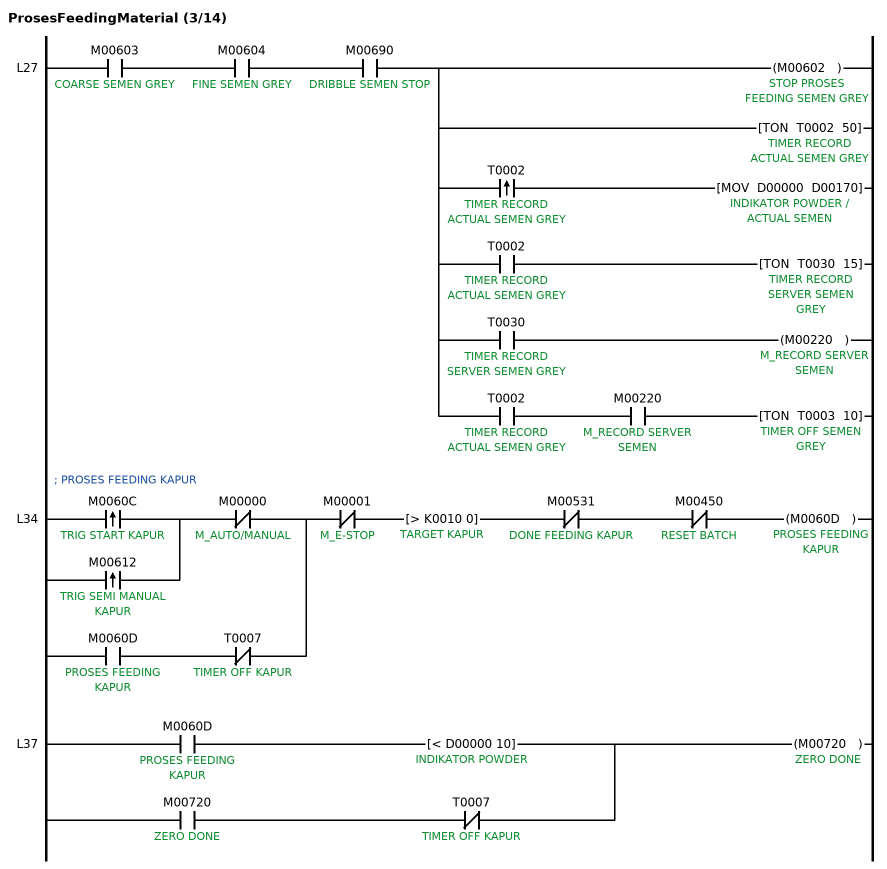
[picture p24: ProsesFeedingMaterial rungs L27-L37]
; L27
LOAD      M00603	// COARSE SEMEN GREY
AND       M00604	// FINE SEMEN GREY
AND       M00690	// DRIBBLE SEMEN STOP
OUT       M00602	// STOP PROSES FEEDING SEMEN GREY 
TON       T0002 50	// TIMER RECORD ACTUAL SEMEN GREY 
MPUSH
ANDP      T0002	// TIMER RECORD ACTUAL SEMEN GREY 
MOV       D00000 D00170	// INDIKATOR POWDER / ACTUAL SEMEN
MLOAD
AND       T0002	// TIMER RECORD ACTUAL SEMEN GREY 
TON       T0030 15	// TIMER RECORD SERVER SEMEN GREY
MLOAD
AND       T0030	// TIMER RECORD SERVER SEMEN GREY
OUT       M00220	// M_RECORD SERVER SEMEN
MPOP
AND       T0002	// TIMER RECORD ACTUAL SEMEN GREY 
AND       M00220	// M_RECORD SERVER SEMEN
TON       T0003 10	// TIMER OFF SEMEN GREY 
// PROSES FEEDING KAPUR
; L34
LOADP     M0060C	// TRIG START KAPUR
ORP       M00612	// TRIG SEMI MANUAL KAPUR 
AND NOT   M00000	// M_AUTO/MANUAL
LOAD      M0060D	// PROSES FEEDING KAPUR 
AND NOT   T0007	// TIMER OFF KAPUR
OR LOAD
AND NOT   M00001	// M_E-STOP
AND>      K0010 0	// TARGET KAPUR 
AND NOT   M00531	// DONE FEEDING KAPUR
AND NOT   M00450	// RESET BATCH
OUT       M0060D	// PROSES FEEDING KAPUR 
; L37
LOAD      M0060D	// PROSES FEEDING KAPUR 
AND<      D00000 10	// INDIKATOR POWDER
LOAD      M00720	// ZERO DONE
AND NOT   T0007	// TIMER OFF KAPUR
OR LOAD
OUT       M00720	// ZERO DONE

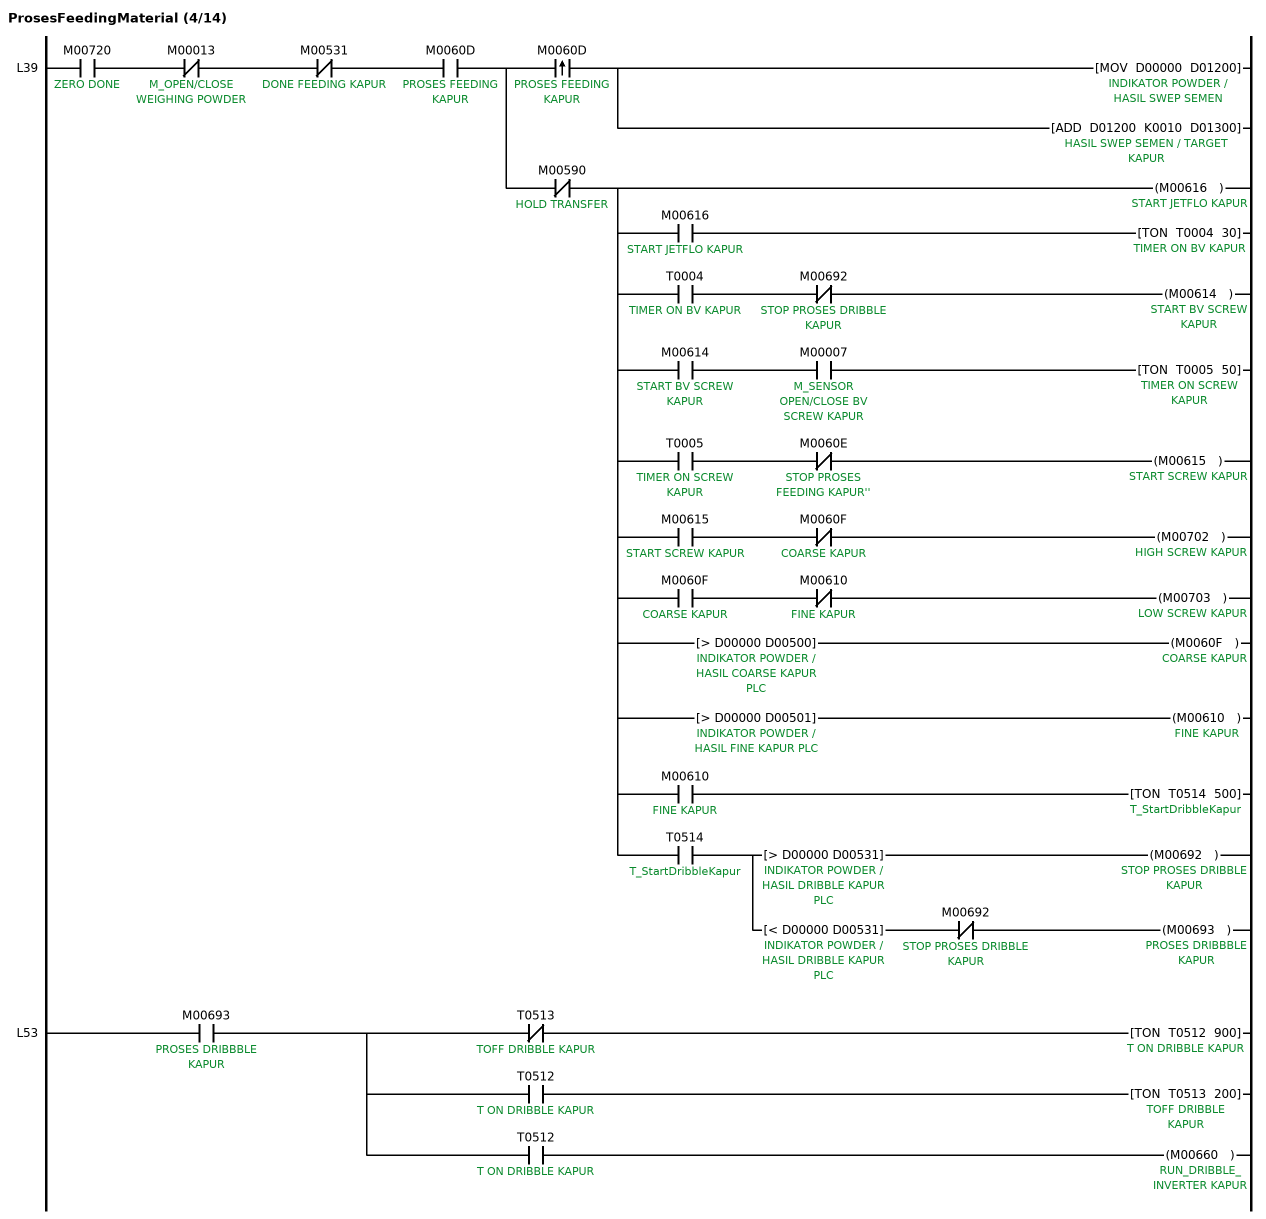
; L39
LOAD      M00720	// ZERO DONE
AND NOT   M00013	// M_OPEN/CLOSE WEIGHING POWDER
AND NOT   M00531	// DONE FEEDING KAPUR
AND       M0060D	// PROSES FEEDING KAPUR 
MPUSH
ANDP      M0060D	// PROSES FEEDING KAPUR 
MOV       D00000 D01200	// INDIKATOR POWDER / HASIL SWEP SEMEN
ADD       D01200 K0010 D01300	// HASIL SWEP SEMEN / TARGET KAPUR 
MPOP
AND NOT   M00590	// HOLD TRANSFER
OUT       M00616	// START JETFLO KAPUR
MPUSH
AND       M00616	// START JETFLO KAPUR
TON       T0004 30	// TIMER ON BV KAPUR
MLOAD
AND       T0004	// TIMER ON BV KAPUR
AND NOT   M00692	// STOP PROSES DRIBBLE KAPUR
OUT       M00614	// START BV SCREW KAPUR
MLOAD
AND       M00614	// START BV SCREW KAPUR
AND       M00007	// M_SENSOR OPEN/CLOSE BV SCREW KAPUR
TON       T0005 50	// TIMER ON SCREW KAPUR
MLOAD
AND       T0005	// TIMER ON SCREW KAPUR
AND NOT   M0060E	// STOP PROSES FEEDING KAPUR''
OUT       M00615	// START SCREW KAPUR
MLOAD
AND       M00615	// START SCREW KAPUR
AND NOT   M0060F	// COARSE KAPUR
OUT       M00702	// HIGH SCREW KAPUR
MLOAD
AND       M0060F	// COARSE KAPUR
AND NOT   M00610	// FINE KAPUR
OUT       M00703	// LOW SCREW KAPUR
MLOAD
AND>      D00000 D00500	// INDIKATOR POWDER / HASIL COARSE KAPUR PLC
OUT       M0060F	// COARSE KAPUR
MLOAD
AND>      D00000 D00501	// INDIKATOR POWDER / HASIL FINE KAPUR PLC 
OUT       M00610	// FINE KAPUR
MLOAD
AND       M00610	// FINE KAPUR
TON       T0514 500	// T_StartDribbleKapur
MPOP
AND       T0514	// T_StartDribbleKapur
MPUSH
AND>      D00000 D00531	// INDIKATOR POWDER / HASIL DRIBBLE KAPUR PLC 
OUT       M00692	// STOP PROSES DRIBBLE KAPUR
MPOP
AND<      D00000 D00531	// INDIKATOR POWDER / HASIL DRIBBLE KAPUR PLC 
AND NOT   M00692	// STOP PROSES DRIBBLE KAPUR
OUT       M00693	// PROSES DRIBBBLE KAPUR
; L53
LOAD      M00693	// PROSES DRIBBBLE KAPUR
MPUSH
AND NOT   T0513	// TOFF DRIBBLE KAPUR
TON       T0512 900	// T ON DRIBBLE KAPUR
MLOAD
AND       T0512	// T ON DRIBBLE KAPUR
TON       T0513 200	// TOFF DRIBBLE KAPUR
MPOP
AND       T0512	// T ON DRIBBLE KAPUR
OUT       M00660	// RUN_DRIBBLE_INVERTER KAPUR

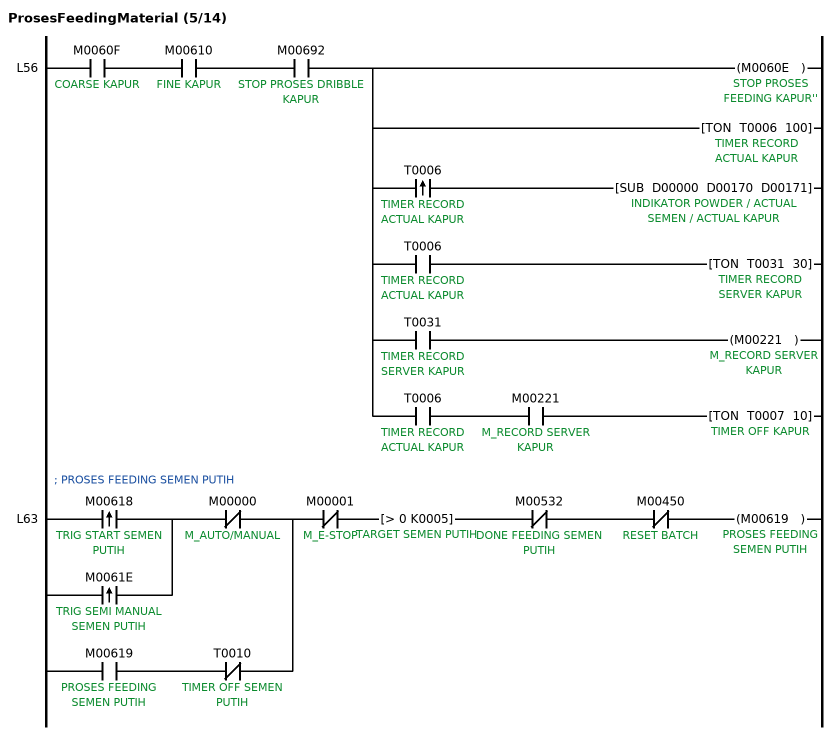
; L56
LOAD      M0060F	// COARSE KAPUR
AND       M00610	// FINE KAPUR
AND       M00692	// STOP PROSES DRIBBLE KAPUR
OUT       M0060E	// STOP PROSES FEEDING KAPUR''
TON       T0006 100	// TIMER RECORD ACTUAL KAPUR
MPUSH
ANDP      T0006	// TIMER RECORD ACTUAL KAPUR
SUB       D00000 D00170 D00171	// INDIKATOR POWDER / ACTUAL SEMEN / ACTUAL KAPUR
MLOAD
AND       T0006	// TIMER RECORD ACTUAL KAPUR
TON       T0031 30	// TIMER RECORD SERVER KAPUR
MLOAD
AND       T0031	// TIMER RECORD SERVER KAPUR
OUT       M00221	// M_RECORD SERVER KAPUR
MPOP
AND       T0006	// TIMER RECORD ACTUAL KAPUR
AND       M00221	// M_RECORD SERVER KAPUR
TON       T0007 10	// TIMER OFF KAPUR
// PROSES FEEDING SEMEN PUTIH
; L63
LOADP     M00618	// TRIG START SEMEN PUTIH
ORP       M0061E	// TRIG SEMI MANUAL SEMEN PUTIH
AND NOT   M00000	// M_AUTO/MANUAL
LOAD      M00619	// PROSES FEEDING SEMEN PUTIH 
AND NOT   T0010	// TIMER OFF SEMEN PUTIH
OR LOAD
AND NOT   M00001	// M_E-STOP
AND>      0 K0005	// TARGET SEMEN PUTIH
AND NOT   M00532	// DONE FEEDING SEMEN PUTIH 
AND NOT   M00450	// RESET BATCH
OUT       M00619	// PROSES FEEDING SEMEN PUTIH 

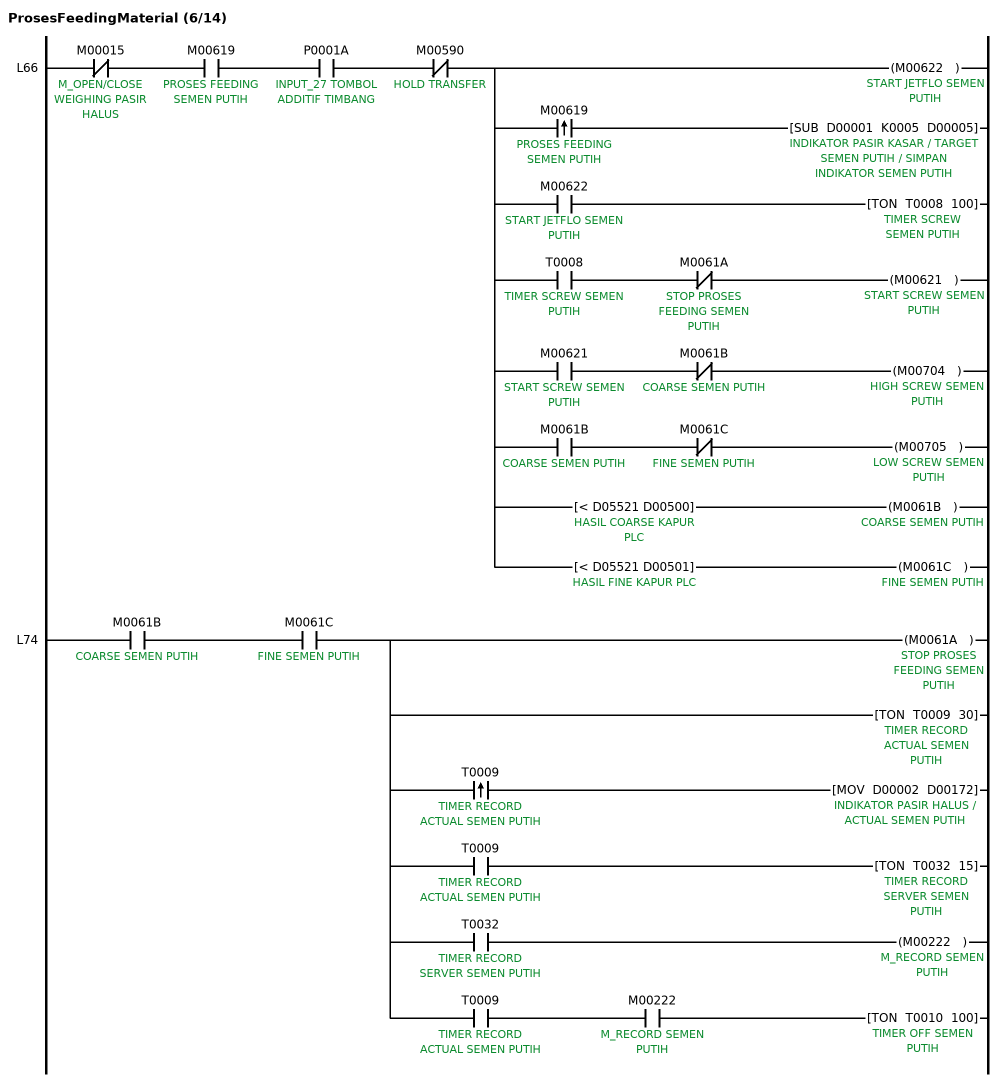
; L66
LOAD NOT  M00015	// M_OPEN/CLOSE WEIGHING PASIR HALUS 
AND       M00619	// PROSES FEEDING SEMEN PUTIH 
AND       P0001A	// INPUT_27 TOMBOL ADDITIF TIMBANG 
AND NOT   M00590	// HOLD TRANSFER
OUT       M00622	// START JETFLO SEMEN PUTIH
MPUSH
ANDP      M00619	// PROSES FEEDING SEMEN PUTIH 
SUB       D00001 K0005 D00005	// INDIKATOR PASIR KASAR / TARGET SEMEN PUTIH / SIMPAN INDIKATOR SEMEN PUTIH 
MLOAD
AND       M00622	// START JETFLO SEMEN PUTIH
TON       T0008 100	// TIMER SCREW SEMEN PUTIH
MLOAD
AND       T0008	// TIMER SCREW SEMEN PUTIH
AND NOT   M0061A	// STOP PROSES FEEDING SEMEN PUTIH
OUT       M00621	// START SCREW SEMEN PUTIH
MLOAD
AND       M00621	// START SCREW SEMEN PUTIH
AND NOT   M0061B	// COARSE SEMEN PUTIH
OUT       M00704	// HIGH SCREW SEMEN PUTIH 
MLOAD
AND       M0061B	// COARSE SEMEN PUTIH
AND NOT   M0061C	// FINE SEMEN PUTIH
OUT       M00705	// LOW SCREW SEMEN PUTIH 
MLOAD
AND<      D05521 D00500	// HASIL COARSE KAPUR PLC
OUT       M0061B	// COARSE SEMEN PUTIH
MPOP
AND<      D05521 D00501	// HASIL FINE KAPUR PLC 
OUT       M0061C	// FINE SEMEN PUTIH
; L74
LOAD      M0061B	// COARSE SEMEN PUTIH
AND       M0061C	// FINE SEMEN PUTIH
OUT       M0061A	// STOP PROSES FEEDING SEMEN PUTIH
TON       T0009 30	// TIMER RECORD ACTUAL SEMEN PUTIH
MPUSH
ANDP      T0009	// TIMER RECORD ACTUAL SEMEN PUTIH
MOV       D00002 D00172	// INDIKATOR PASIR HALUS / ACTUAL SEMEN PUTIH
MLOAD
AND       T0009	// TIMER RECORD ACTUAL SEMEN PUTIH
TON       T0032 15	// TIMER RECORD SERVER SEMEN PUTIH
MLOAD
AND       T0032	// TIMER RECORD SERVER SEMEN PUTIH
OUT       M00222	// M_RECORD SEMEN PUTIH
MPOP
AND       T0009	// TIMER RECORD ACTUAL SEMEN PUTIH
AND       M00222	// M_RECORD SEMEN PUTIH
TON       T0010 100	// TIMER OFF SEMEN PUTIH

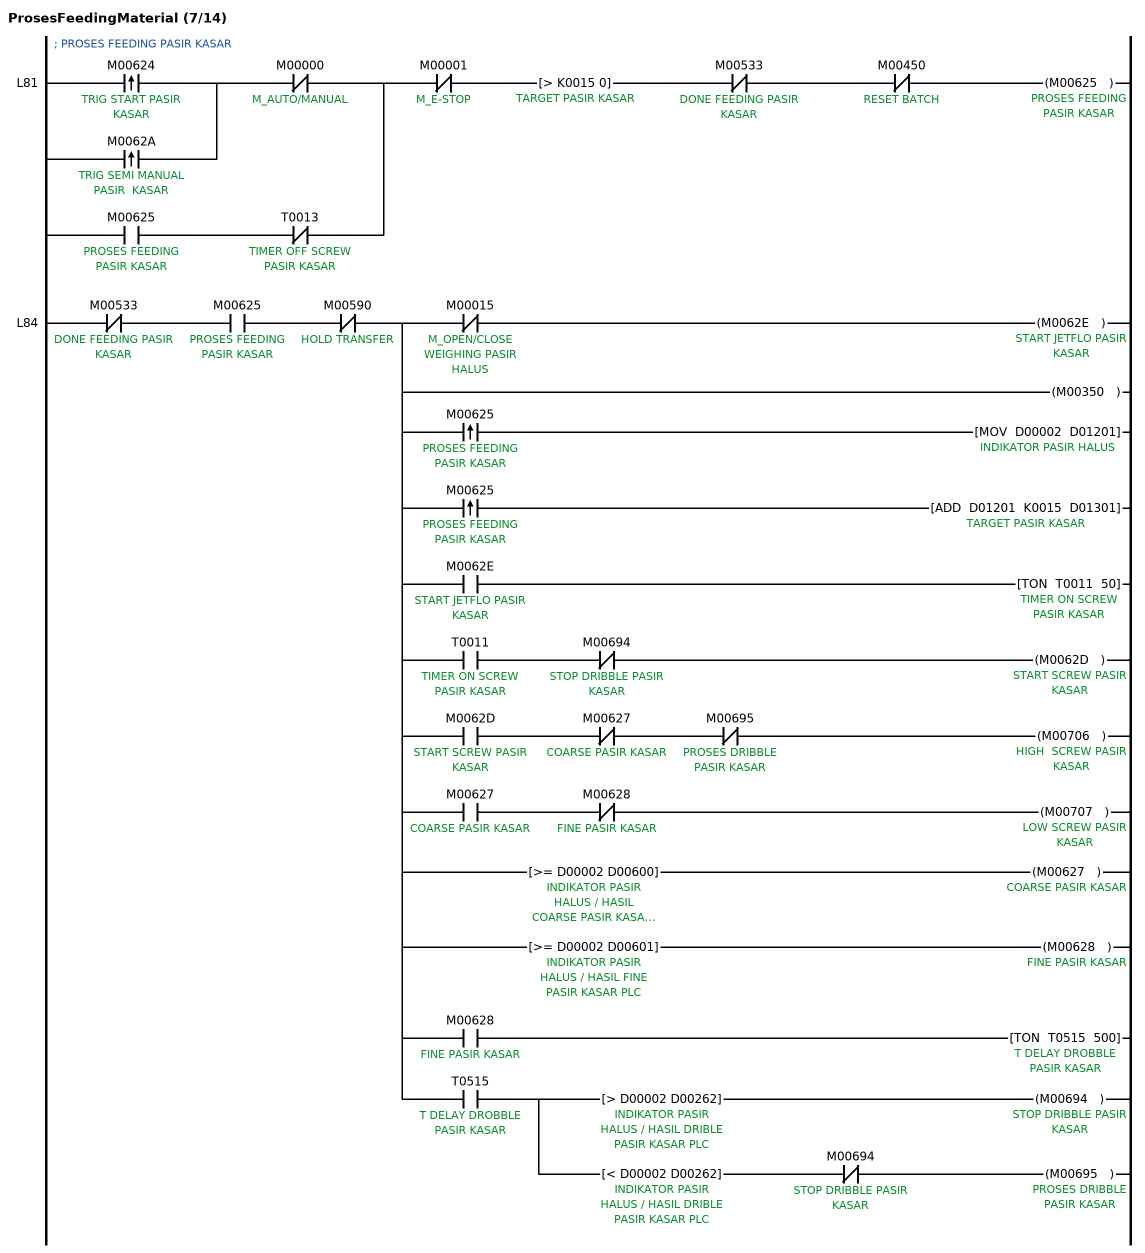
// PROSES FEEDING PASIR KASAR
; L81
LOADP     M00624	// TRIG START PASIR KASAR
ORP       M0062A	// TRIG SEMI MANUAL PASIR  KASAR
AND NOT   M00000	// M_AUTO/MANUAL
LOAD      M00625	// PROSES FEEDING PASIR KASAR
AND NOT   T0013	// TIMER OFF SCREW PASIR KASAR
OR LOAD
AND NOT   M00001	// M_E-STOP
AND>      K0015 0	// TARGET PASIR KASAR
AND NOT   M00533	// DONE FEEDING PASIR KASAR
AND NOT   M00450	// RESET BATCH
OUT       M00625	// PROSES FEEDING PASIR KASAR
; L84
LOAD NOT  M00533	// DONE FEEDING PASIR KASAR
AND       M00625	// PROSES FEEDING PASIR KASAR
AND NOT   M00590	// HOLD TRANSFER
MPUSH
AND NOT   M00015	// M_OPEN/CLOSE WEIGHING PASIR HALUS 
OUT       M0062E	// START JETFLO PASIR KASAR
MLOAD
OUT       M00350
ANDP      M00625	// PROSES FEEDING PASIR KASAR
MOV       D00002 D01201	// INDIKATOR PASIR HALUS
MLOAD
ANDP      M00625	// PROSES FEEDING PASIR KASAR
ADD       D01201 K0015 D01301	// TARGET PASIR KASAR
MLOAD
AND       M0062E	// START JETFLO PASIR KASAR
TON       T0011 50	// TIMER ON SCREW PASIR KASAR
MLOAD
AND       T0011	// TIMER ON SCREW PASIR KASAR
AND NOT   M00694	// STOP DRIBBLE PASIR KASAR
OUT       M0062D	// START SCREW PASIR KASAR
MLOAD
AND       M0062D	// START SCREW PASIR KASAR
AND NOT   M00627	// COARSE PASIR KASAR
AND NOT   M00695	// PROSES DRIBBLE PASIR KASAR
OUT       M00706	// HIGH  SCREW PASIR KASAR
MLOAD
AND       M00627	// COARSE PASIR KASAR
AND NOT   M00628	// FINE PASIR KASAR
OUT       M00707	// LOW SCREW PASIR KASAR
MLOAD
AND>=     D00002 D00600	// INDIKATOR PASIR HALUS / HASIL COARSE PASIR KASAR PLC
OUT       M00627	// COARSE PASIR KASAR
MLOAD
AND>=     D00002 D00601	// INDIKATOR PASIR HALUS / HASIL FINE PASIR KASAR PLC
OUT       M00628	// FINE PASIR KASAR
MLOAD
AND       M00628	// FINE PASIR KASAR
TON       T0515 500	// T DELAY DROBBLE PASIR KASAR
MPOP
AND       T0515	// T DELAY DROBBLE PASIR KASAR
MPUSH
AND>      D00002 D00262	// INDIKATOR PASIR HALUS / HASIL DRIBLE PASIR KASAR PLC
OUT       M00694	// STOP DRIBBLE PASIR KASAR
MPOP
AND<      D00002 D00262	// INDIKATOR PASIR HALUS / HASIL DRIBLE PASIR KASAR PLC
AND NOT   M00694	// STOP DRIBBLE PASIR KASAR
OUT       M00695	// PROSES DRIBBLE PASIR KASAR

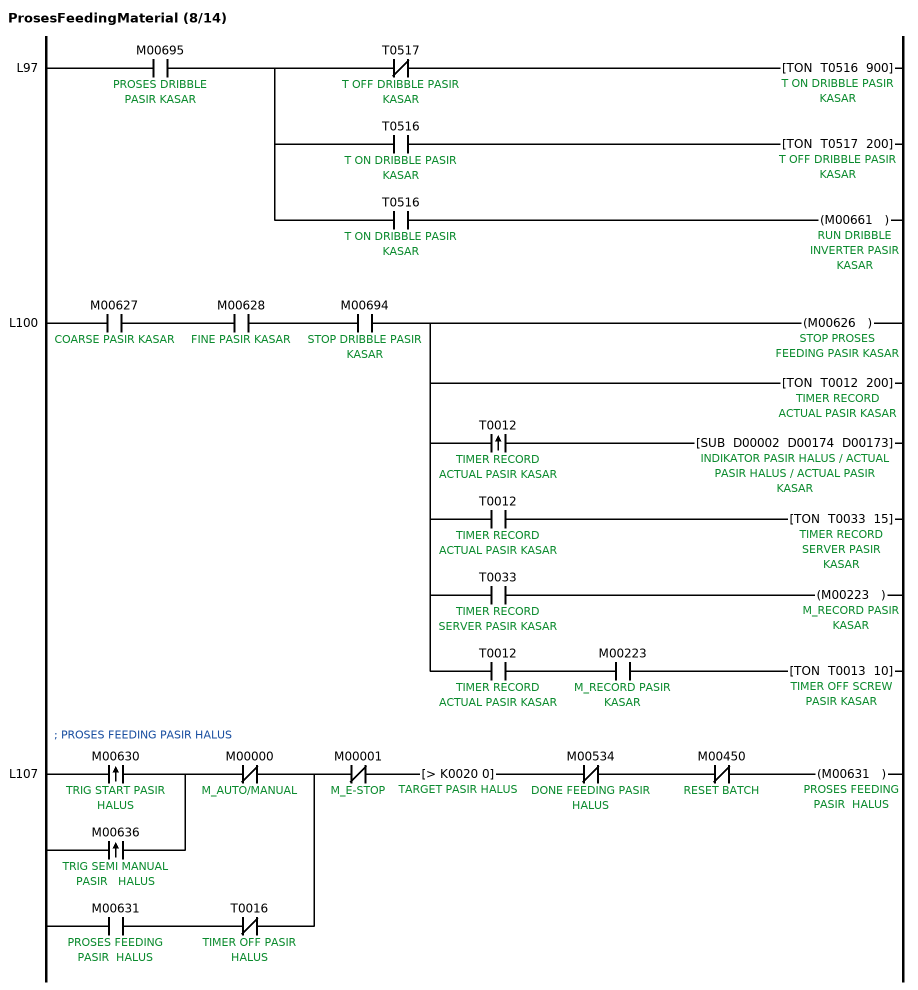
; L97
LOAD      M00695	// PROSES DRIBBLE PASIR KASAR
MPUSH
AND NOT   T0517	// T OFF DRIBBLE PASIR KASAR
TON       T0516 900	// T ON DRIBBLE PASIR KASAR
MLOAD
AND       T0516	// T ON DRIBBLE PASIR KASAR
TON       T0517 200	// T OFF DRIBBLE PASIR KASAR
MPOP
AND       T0516	// T ON DRIBBLE PASIR KASAR
OUT       M00661	// RUN DRIBBLE INVERTER PASIR KASAR
; L100
LOAD      M00627	// COARSE PASIR KASAR
AND       M00628	// FINE PASIR KASAR
AND       M00694	// STOP DRIBBLE PASIR KASAR
OUT       M00626	// STOP PROSES FEEDING PASIR KASAR
TON       T0012 200	// TIMER RECORD ACTUAL PASIR KASAR
MPUSH
ANDP      T0012	// TIMER RECORD ACTUAL PASIR KASAR
SUB       D00002 D00174 D00173	// INDIKATOR PASIR HALUS / ACTUAL PASIR HALUS / ACTUAL PASIR KASAR
MLOAD
AND       T0012	// TIMER RECORD ACTUAL PASIR KASAR
TON       T0033 15	// TIMER RECORD SERVER PASIR KASAR
MLOAD
AND       T0033	// TIMER RECORD SERVER PASIR KASAR
OUT       M00223	// M_RECORD PASIR KASAR
MPOP
AND       T0012	// TIMER RECORD ACTUAL PASIR KASAR
AND       M00223	// M_RECORD PASIR KASAR
TON       T0013 10	// TIMER OFF SCREW PASIR KASAR
// PROSES FEEDING PASIR HALUS
; L107
LOADP     M00630	// TRIG START PASIR HALUS
ORP       M00636	// TRIG SEMI MANUAL PASIR   HALUS
AND NOT   M00000	// M_AUTO/MANUAL
LOAD      M00631	// PROSES FEEDING PASIR  HALUS
AND NOT   T0016	// TIMER OFF PASIR HALUS 
OR LOAD
AND NOT   M00001	// M_E-STOP
AND>      K0020 0	// TARGET PASIR HALUS 
AND NOT   M00534	// DONE FEEDING PASIR HALUS
AND NOT   M00450	// RESET BATCH
OUT       M00631	// PROSES FEEDING PASIR  HALUS

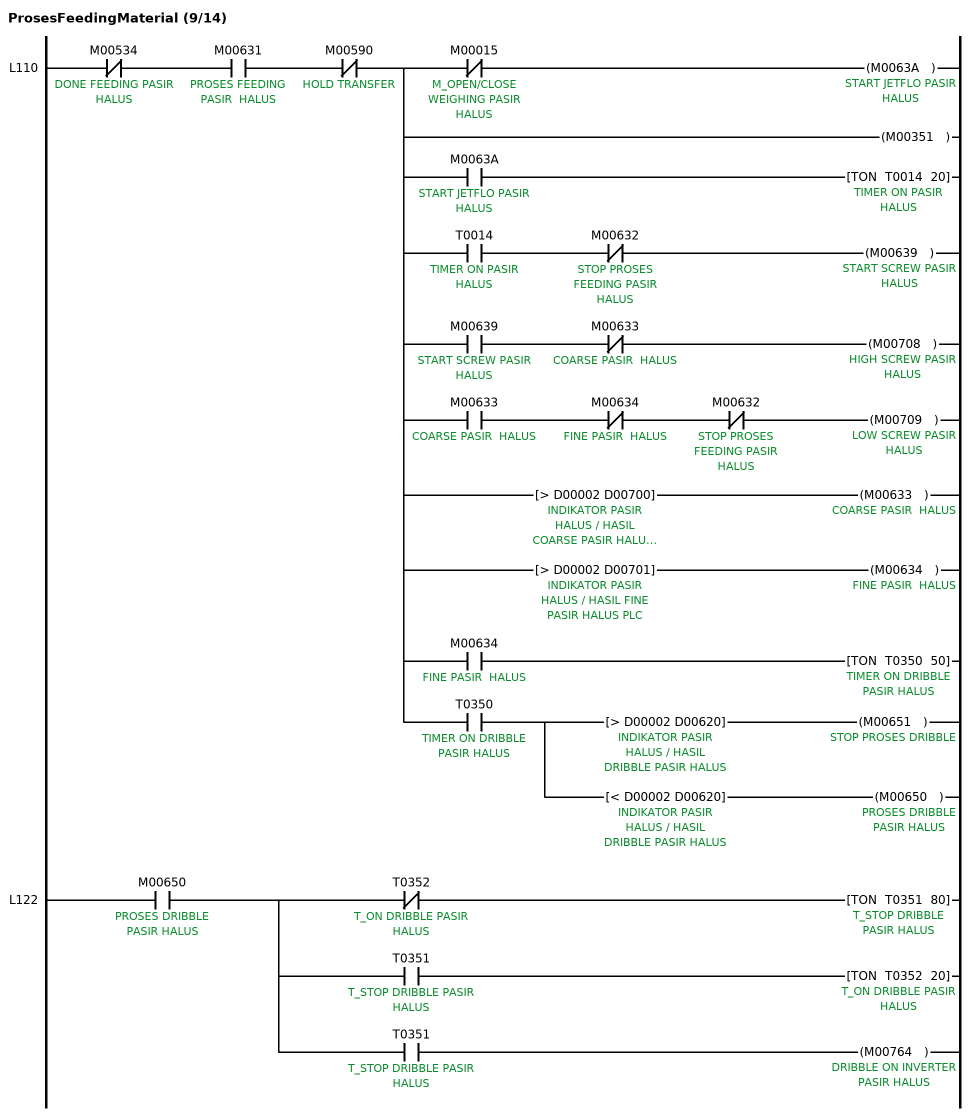
; L110
LOAD NOT  M00534	// DONE FEEDING PASIR HALUS
AND       M00631	// PROSES FEEDING PASIR  HALUS
AND NOT   M00590	// HOLD TRANSFER
MPUSH
AND NOT   M00015	// M_OPEN/CLOSE WEIGHING PASIR HALUS 
OUT       M0063A	// START JETFLO PASIR  HALUS
MLOAD
OUT       M00351
AND       M0063A	// START JETFLO PASIR  HALUS
TON       T0014 20	// TIMER ON PASIR HALUS 
MLOAD
AND       T0014	// TIMER ON PASIR HALUS 
AND NOT   M00632	// STOP PROSES FEEDING PASIR  HALUS
OUT       M00639	// START SCREW PASIR  HALUS
MLOAD
AND       M00639	// START SCREW PASIR  HALUS
AND NOT   M00633	// COARSE PASIR  HALUS
OUT       M00708	// HIGH SCREW PASIR HALUS
MLOAD
AND       M00633	// COARSE PASIR  HALUS
AND NOT   M00634	// FINE PASIR  HALUS
AND NOT   M00632	// STOP PROSES FEEDING PASIR  HALUS
OUT       M00709	// LOW SCREW PASIR HALUS 
MLOAD
AND>      D00002 D00700	// INDIKATOR PASIR HALUS / HASIL COARSE PASIR HALUS PLC
OUT       M00633	// COARSE PASIR  HALUS
MLOAD
AND>      D00002 D00701	// INDIKATOR PASIR HALUS / HASIL FINE PASIR HALUS PLC
OUT       M00634	// FINE PASIR  HALUS
MLOAD
AND       M00634	// FINE PASIR  HALUS
TON       T0350 50	// TIMER ON DRIBBLE PASIR HALUS
MPOP
AND       T0350	// TIMER ON DRIBBLE PASIR HALUS
MPUSH
AND>      D00002 D00620	// INDIKATOR PASIR HALUS / HASIL DRIBBLE PASIR HALUS
OUT       M00651	// STOP PROSES DRIBBLE
MPOP
AND<      D00002 D00620	// INDIKATOR PASIR HALUS / HASIL DRIBBLE PASIR HALUS
OUT       M00650	// PROSES DRIBBLE PASIR HALUS
; L122
LOAD      M00650	// PROSES DRIBBLE PASIR HALUS
MPUSH
AND NOT   T0352	// T_ON DRIBBLE PASIR HALUS
TON       T0351 80	// T_STOP DRIBBLE PASIR HALUS
MLOAD
AND       T0351	// T_STOP DRIBBLE PASIR HALUS
TON       T0352 20	// T_ON DRIBBLE PASIR HALUS
MPOP
AND       T0351	// T_STOP DRIBBLE PASIR HALUS
OUT       M00764	// DRIBBLE ON INVERTER PASIR HALUS

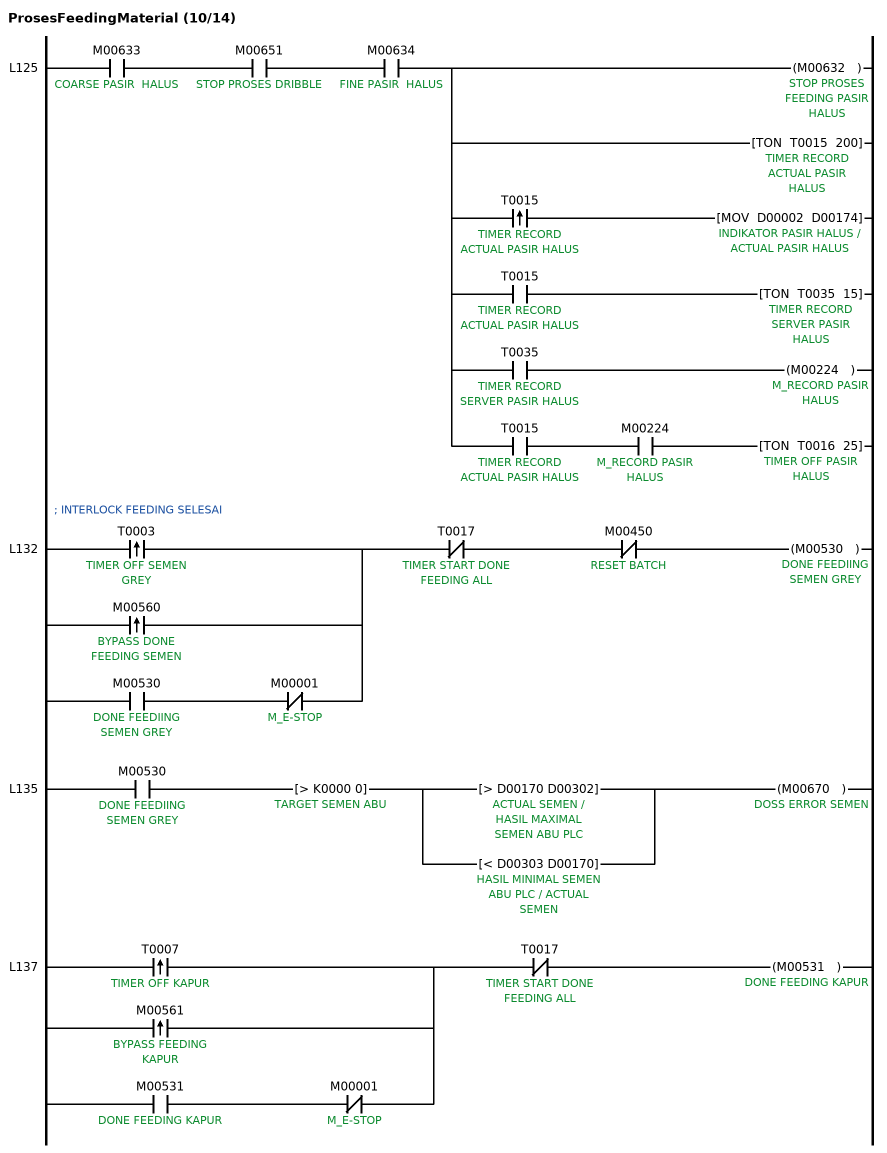
; L125
LOAD      M00633	// COARSE PASIR  HALUS
AND       M00651	// STOP PROSES DRIBBLE
AND       M00634	// FINE PASIR  HALUS
OUT       M00632	// STOP PROSES FEEDING PASIR  HALUS
TON       T0015 200	// TIMER RECORD ACTUAL PASIR HALUS 
MPUSH
ANDP      T0015	// TIMER RECORD ACTUAL PASIR HALUS 
MOV       D00002 D00174	// INDIKATOR PASIR HALUS / ACTUAL PASIR HALUS
MLOAD
AND       T0015	// TIMER RECORD ACTUAL PASIR HALUS 
TON       T0035 15	// TIMER RECORD SERVER PASIR HALUS
MLOAD
AND       T0035	// TIMER RECORD SERVER PASIR HALUS
OUT       M00224	// M_RECORD PASIR HALUS
MPOP
AND       T0015	// TIMER RECORD ACTUAL PASIR HALUS 
AND       M00224	// M_RECORD PASIR HALUS
TON       T0016 25	// TIMER OFF PASIR HALUS 
// INTERLOCK FEEDING SELESAI
; L132
LOADP     T0003	// TIMER OFF SEMEN GREY 
ORP       M00560	// BYPASS DONE FEEDING SEMEN
LOAD      M00530	// DONE FEEDIING SEMEN GREY 
AND NOT   M00001	// M_E-STOP
OR LOAD
AND NOT   T0017	// TIMER START DONE FEEDING ALL 
AND NOT   M00450	// RESET BATCH
OUT       M00530	// DONE FEEDIING SEMEN GREY 
; L135
LOAD      M00530	// DONE FEEDIING SEMEN GREY 
AND>      K0000 0	// TARGET SEMEN ABU 
LOAD>     D00170 D00302	// ACTUAL SEMEN / HASIL MAXIMAL SEMEN ABU PLC
OR<       D00303 D00170	// HASIL MINIMAL SEMEN ABU PLC / ACTUAL SEMEN
AND LOAD
OUT       M00670	// DOSS ERROR SEMEN
; L137
LOADP     T0007	// TIMER OFF KAPUR
ORP       M00561	// BYPASS FEEDING KAPUR
LOAD      M00531	// DONE FEEDING KAPUR
AND NOT   M00001	// M_E-STOP
OR LOAD
AND NOT   T0017	// TIMER START DONE FEEDING ALL 
OUT       M00531	// DONE FEEDING KAPUR

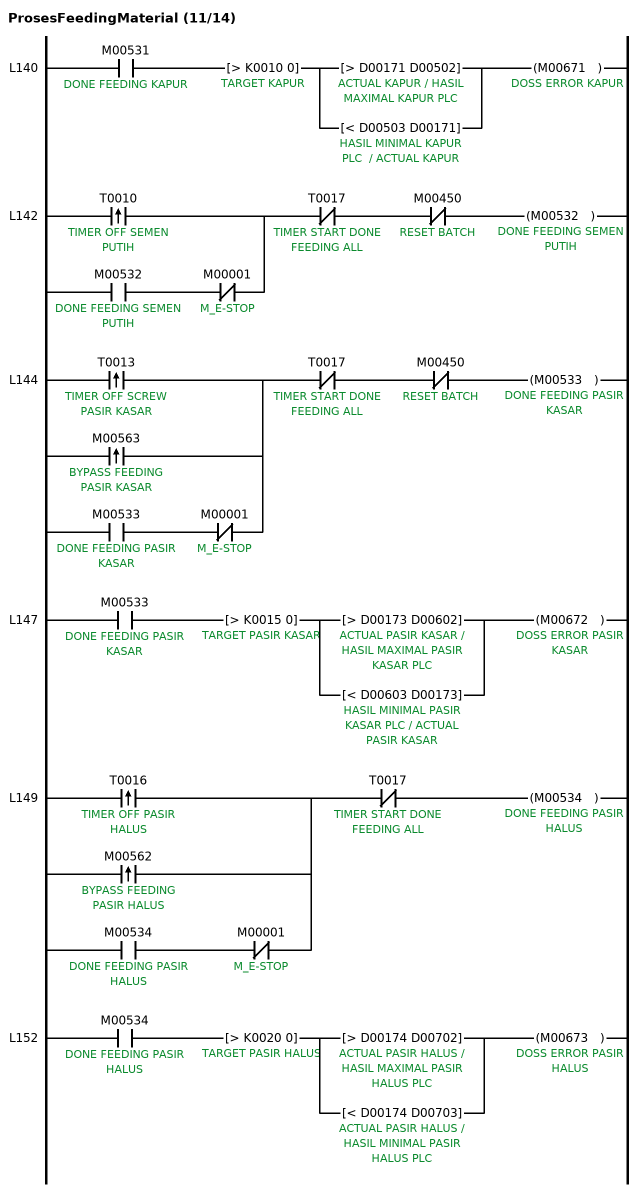
; L140
LOAD      M00531	// DONE FEEDING KAPUR
AND>      K0010 0	// TARGET KAPUR 
LOAD>     D00171 D00502	// ACTUAL KAPUR / HASIL MAXIMAL KAPUR PLC 
OR<       D00503 D00171	// HASIL MINIMAL KAPUR PLC  / ACTUAL KAPUR
AND LOAD
OUT       M00671	// DOSS ERROR KAPUR
; L142
LOADP     T0010	// TIMER OFF SEMEN PUTIH
LOAD      M00532	// DONE FEEDING SEMEN PUTIH 
AND NOT   M00001	// M_E-STOP
OR LOAD
AND NOT   T0017	// TIMER START DONE FEEDING ALL 
AND NOT   M00450	// RESET BATCH
OUT       M00532	// DONE FEEDING SEMEN PUTIH 
; L144
LOADP     T0013	// TIMER OFF SCREW PASIR KASAR
ORP       M00563	// BYPASS FEEDING PASIR KASAR
LOAD      M00533	// DONE FEEDING PASIR KASAR
AND NOT   M00001	// M_E-STOP
OR LOAD
AND NOT   T0017	// TIMER START DONE FEEDING ALL 
AND NOT   M00450	// RESET BATCH
OUT       M00533	// DONE FEEDING PASIR KASAR
; L147
LOAD      M00533	// DONE FEEDING PASIR KASAR
AND>      K0015 0	// TARGET PASIR KASAR
LOAD>     D00173 D00602	// ACTUAL PASIR KASAR / HASIL MAXIMAL PASIR KASAR PLC
OR<       D00603 D00173	// HASIL MINIMAL PASIR KASAR PLC / ACTUAL PASIR KASAR
AND LOAD
OUT       M00672	// DOSS ERROR PASIR KASAR
; L149
LOADP     T0016	// TIMER OFF PASIR HALUS 
ORP       M00562	// BYPASS FEEDING PASIR HALUS
LOAD      M00534	// DONE FEEDING PASIR HALUS
AND NOT   M00001	// M_E-STOP
OR LOAD
AND NOT   T0017	// TIMER START DONE FEEDING ALL 
OUT       M00534	// DONE FEEDING PASIR HALUS
; L152
LOAD      M00534	// DONE FEEDING PASIR HALUS
AND>      K0020 0	// TARGET PASIR HALUS 
LOAD>     D00174 D00702	// ACTUAL PASIR HALUS / HASIL MAXIMAL PASIR HALUS PLC
OR<       D00174 D00703	// ACTUAL PASIR HALUS / HASIL MINIMAL PASIR HALUS PLC
AND LOAD
OUT       M00673	// DOSS ERROR PASIR HALUS

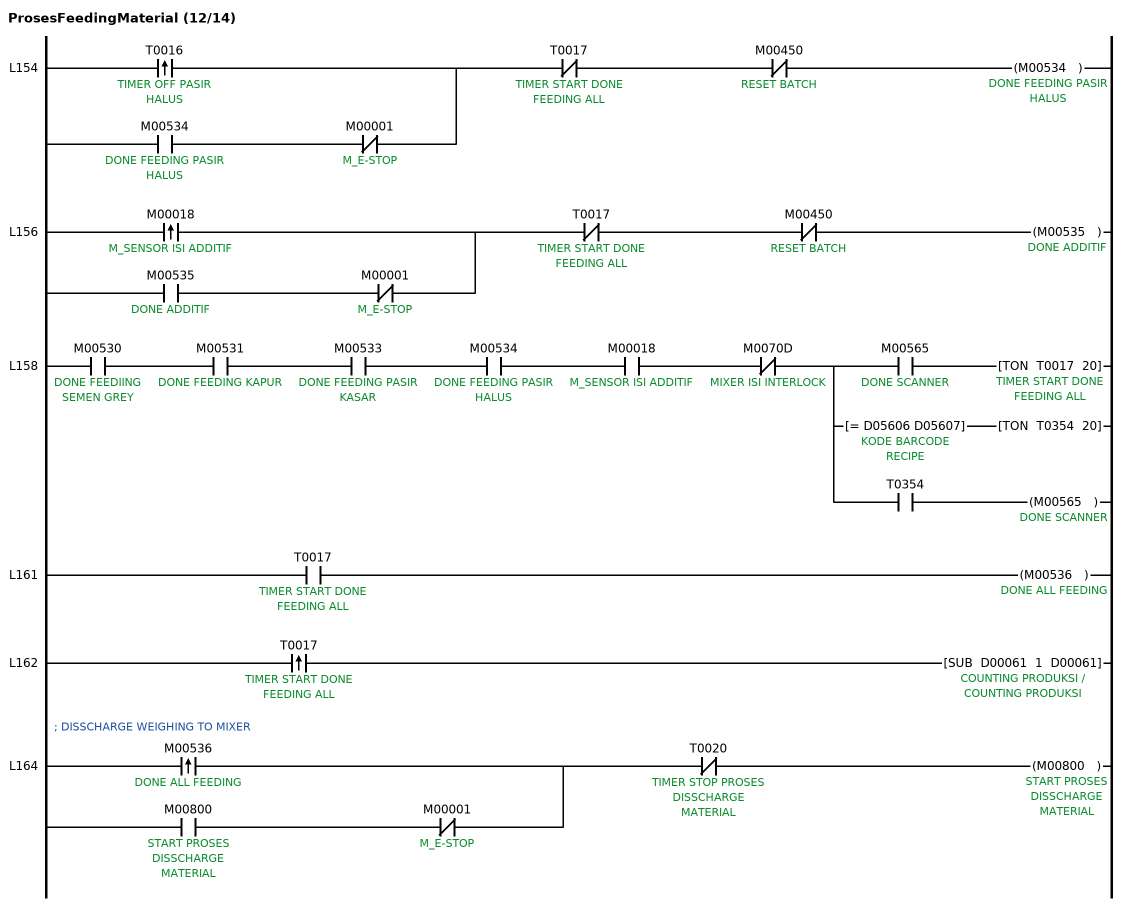
; L154
LOADP     T0016	// TIMER OFF PASIR HALUS 
LOAD      M00534	// DONE FEEDING PASIR HALUS
AND NOT   M00001	// M_E-STOP
OR LOAD
AND NOT   T0017	// TIMER START DONE FEEDING ALL 
AND NOT   M00450	// RESET BATCH
OUT       M00534	// DONE FEEDING PASIR HALUS
; L156
LOADP     M00018	// M_SENSOR ISI ADDITIF
LOAD      M00535	// DONE ADDITIF 
AND NOT   M00001	// M_E-STOP
OR LOAD
AND NOT   T0017	// TIMER START DONE FEEDING ALL 
AND NOT   M00450	// RESET BATCH
OUT       M00535	// DONE ADDITIF 
; L158
LOAD      M00530	// DONE FEEDIING SEMEN GREY 
AND       M00531	// DONE FEEDING KAPUR
AND       M00533	// DONE FEEDING PASIR KASAR
AND       M00534	// DONE FEEDING PASIR HALUS
AND       M00018	// M_SENSOR ISI ADDITIF
AND NOT   M0070D	// MIXER ISI INTERLOCK
MPUSH
AND       M00565	// DONE SCANNER
TON       T0017 20	// TIMER START DONE FEEDING ALL 
MLOAD
AND=      D05606 D05607	// KODE BARCODE RECIPE
TON       T0354 20
MPOP
AND       T0354
OUT       M00565	// DONE SCANNER
; L161
LOAD      T0017	// TIMER START DONE FEEDING ALL 
OUT       M00536	// DONE ALL FEEDING 
; L162
LOADP     T0017	// TIMER START DONE FEEDING ALL 
SUB       D00061 1 D00061	// COUNTING PRODUKSI / COUNTING PRODUKSI
// DISSCHARGE WEIGHING TO MIXER
; L164
LOADP     M00536	// DONE ALL FEEDING 
LOAD      M00800	// START PROSES DISSCHARGE MATERIAL 
AND NOT   M00001	// M_E-STOP
OR LOAD
AND NOT   T0020	// TIMER STOP PROSES DISSCHARGE MATERIAL 
OUT       M00800	// START PROSES DISSCHARGE MATERIAL 

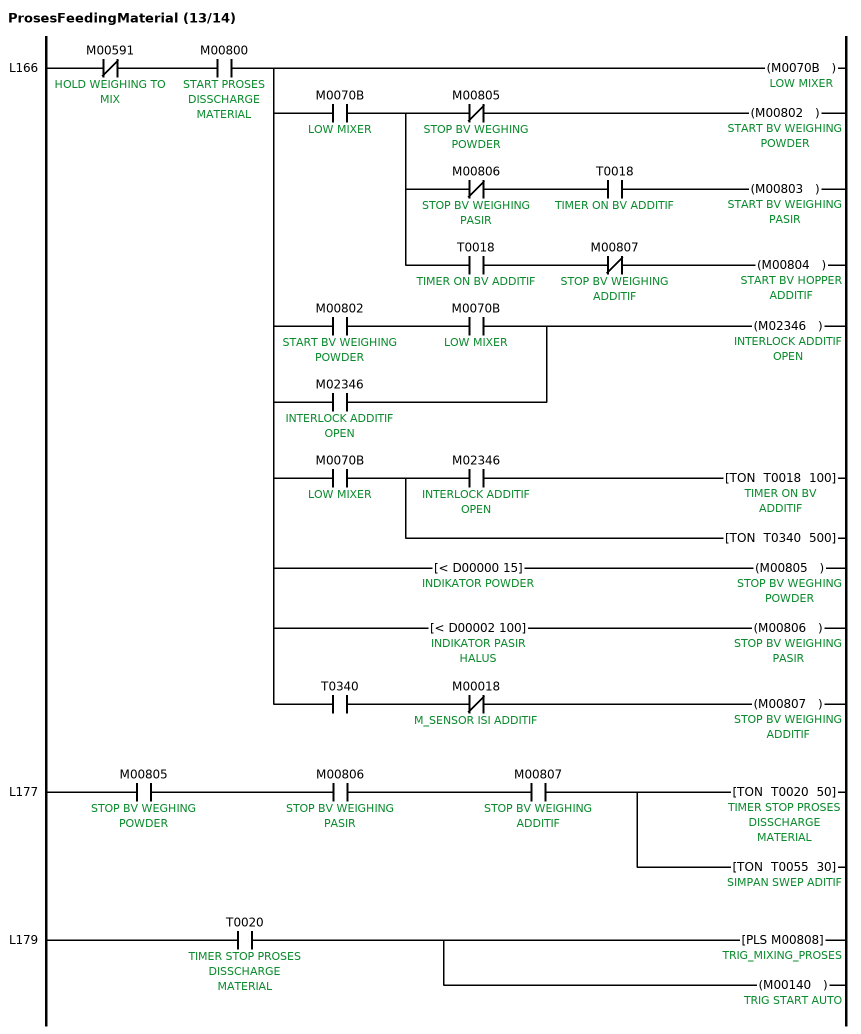
; L166
LOAD NOT  M00591	// HOLD WEIGHING TO MIX
AND       M00800	// START PROSES DISSCHARGE MATERIAL 
OUT       M0070B	// LOW MIXER 
MPUSH
AND       M0070B	// LOW MIXER 
MPUSH
AND NOT   M00805	// STOP BV WEGHING  POWDER 
OUT       M00802	// START BV WEIGHING POWDER 
MLOAD
AND NOT   M00806	// STOP BV WEIGHING PASIR
AND       T0018	// TIMER ON BV ADDITIF 
OUT       M00803	// START BV WEIGHING PASIR 
MPOP
AND       T0018	// TIMER ON BV ADDITIF 
AND NOT   M00807	// STOP BV WEIGHING ADDITIF
OUT       M00804	// START BV HOPPER ADDITIF 
MLOAD
LOAD      M00802	// START BV WEIGHING POWDER 
AND       M0070B	// LOW MIXER 
OR        M02346	// INTERLOCK ADDITIF OPEN
AND LOAD
OUT       M02346	// INTERLOCK ADDITIF OPEN
MLOAD
AND       M0070B	// LOW MIXER 
MPUSH
AND       M02346	// INTERLOCK ADDITIF OPEN
TON       T0018 100	// TIMER ON BV ADDITIF 
MPOP
TON       T0340 500
MLOAD
AND<      D00000 15	// INDIKATOR POWDER
OUT       M00805	// STOP BV WEGHING  POWDER 
MLOAD
AND<      D00002 100	// INDIKATOR PASIR HALUS
OUT       M00806	// STOP BV WEIGHING PASIR
MPOP
AND       T0340
AND NOT   M00018	// M_SENSOR ISI ADDITIF
OUT       M00807	// STOP BV WEIGHING ADDITIF
; L177
LOAD      M00805	// STOP BV WEGHING  POWDER 
AND       M00806	// STOP BV WEIGHING PASIR
AND       M00807	// STOP BV WEIGHING ADDITIF
TON       T0020 50	// TIMER STOP PROSES DISSCHARGE MATERIAL 
TON       T0055 30	// SIMPAN SWEP ADITIF
; L179
LOAD      T0020	// TIMER STOP PROSES DISSCHARGE MATERIAL 
OUTP      M00808	// TRIG_MIXING_PROSES
OUT       M00140	// TRIG START AUTO

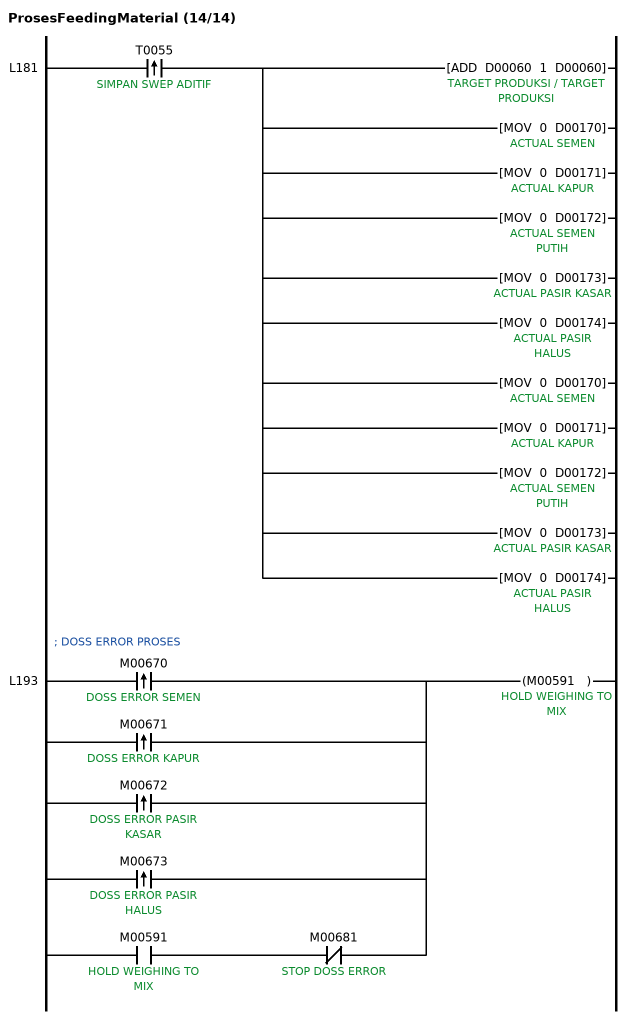
; L181
LOADP     T0055	// SIMPAN SWEP ADITIF
ADD       D00060 1 D00060	// TARGET PRODUKSI / TARGET PRODUKSI
MOV       0 D00170	// ACTUAL SEMEN
MOV       0 D00171	// ACTUAL KAPUR
MOV       0 D00172	// ACTUAL SEMEN PUTIH
MOV       0 D00173	// ACTUAL PASIR KASAR
MOV       0 D00174	// ACTUAL PASIR HALUS
MOV       0 D00170	// ACTUAL SEMEN
MOV       0 D00171	// ACTUAL KAPUR
MOV       0 D00172	// ACTUAL SEMEN PUTIH
MOV       0 D00173	// ACTUAL PASIR KASAR
MOV       0 D00174	// ACTUAL PASIR HALUS
// DOSS ERROR PROSES
; L193
LOADP     M00670	// DOSS ERROR SEMEN
ORP       M00671	// DOSS ERROR KAPUR
ORP       M00672	// DOSS ERROR PASIR KASAR
ORP       M00673	// DOSS ERROR PASIR HALUS
LOAD      M00591	// HOLD WEIGHING TO MIX
AND NOT   M00681	// STOP DOSS ERROR
OR LOAD
OUT       M00591	// HOLD WEIGHING TO MIX

PROGRAM MixingProsesDanDisschargemixProses (task: Scan Program)

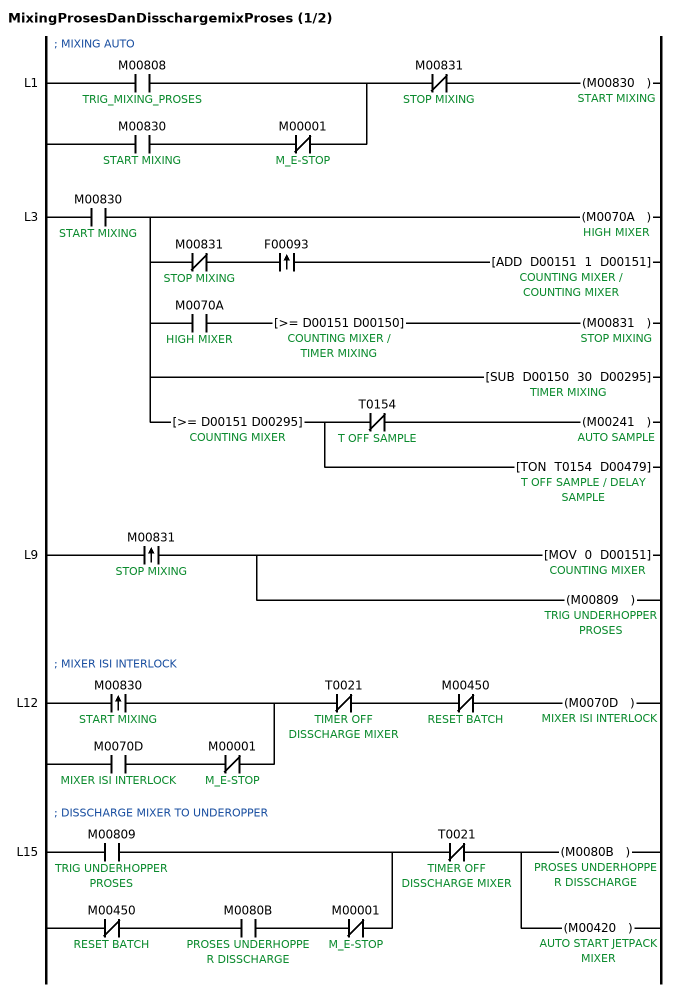
// MIXING AUTO
; L1
LOAD      M00808	// TRIG_MIXING_PROSES
LOAD      M00830	// START MIXING 
AND NOT   M00001	// M_E-STOP
OR LOAD
AND NOT   M00831	// STOP MIXING 
OUT       M00830	// START MIXING 
; L3
LOAD      M00830	// START MIXING 
OUT       M0070A	// HIGH MIXER 
MPUSH
AND NOT   M00831	// STOP MIXING 
ANDP      F00093
ADD       D00151 1 D00151	// COUNTING MIXER / COUNTING MIXER
MLOAD
AND       M0070A	// HIGH MIXER 
AND>=     D00151 D00150	// COUNTING MIXER / TIMER MIXING
OUT       M00831	// STOP MIXING 
MPOP
SUB       D00150 30 D00295	// TIMER MIXING
AND>=     D00151 D00295	// COUNTING MIXER
MPUSH
AND NOT   T0154	// T OFF SAMPLE
OUT       M00241	// AUTO SAMPLE
MPOP
TON       T0154 D00479	// T OFF SAMPLE / DELAY SAMPLE
; L9
LOADP     M00831	// STOP MIXING 
MOV       0 D00151	// COUNTING MIXER
OUT       M00809	// TRIG UNDERHOPPER PROSES 
// MIXER ISI INTERLOCK
; L12
LOADP     M00830	// START MIXING 
LOAD      M0070D	// MIXER ISI INTERLOCK
AND NOT   M00001	// M_E-STOP
OR LOAD
AND NOT   T0021	// TIMER OFF DISSCHARGE MIXER
AND NOT   M00450	// RESET BATCH
OUT       M0070D	// MIXER ISI INTERLOCK
// DISSCHARGE MIXER TO UNDEROPPER
; L15
LOAD      M00809	// TRIG UNDERHOPPER PROSES 
LOAD NOT  M00450	// RESET BATCH
AND       M0080B	// PROSES UNDERHOPPER DISSCHARGE
AND NOT   M00001	// M_E-STOP
OR LOAD
AND NOT   T0021	// TIMER OFF DISSCHARGE MIXER
OUT       M0080B	// PROSES UNDERHOPPER DISSCHARGE
OUT       M00420	// AUTO START JETPACK  MIXER

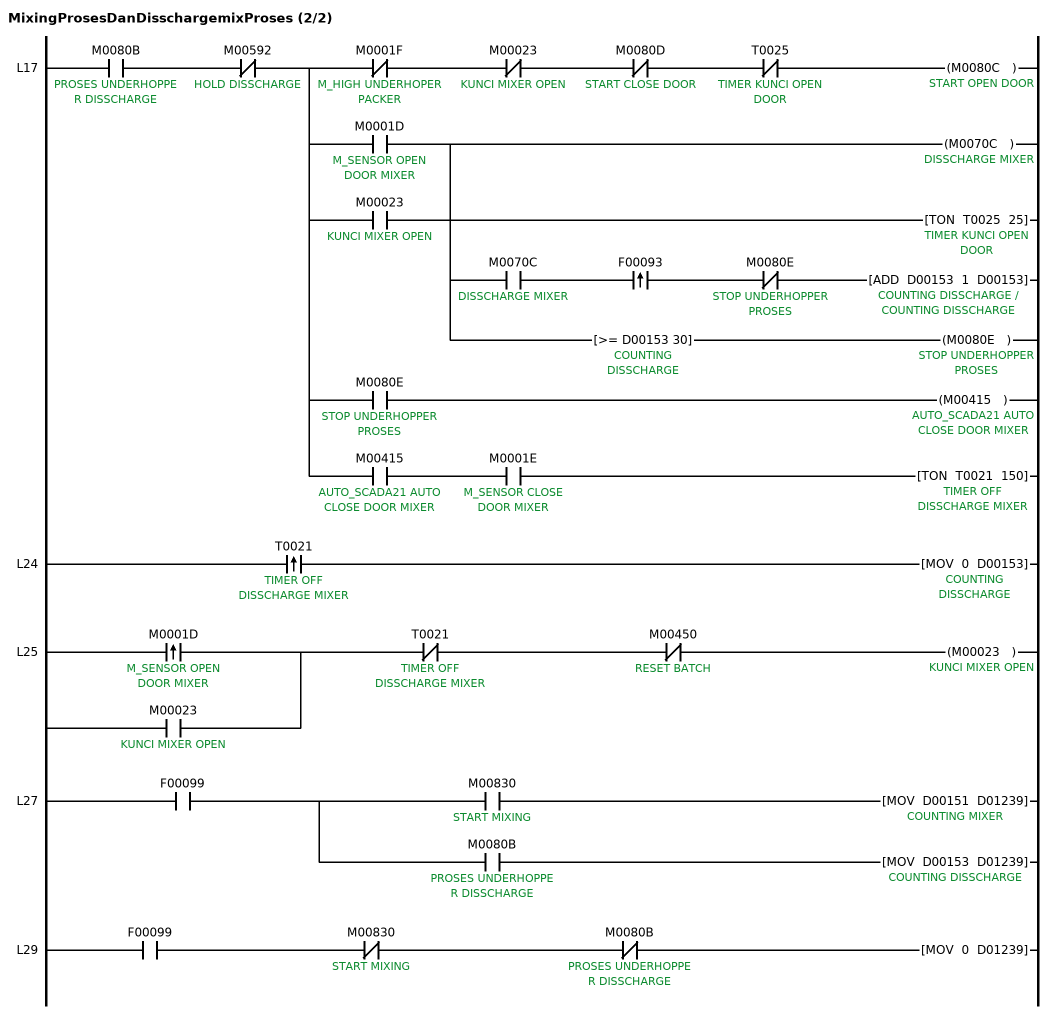
; L17
LOAD      M0080B	// PROSES UNDERHOPPER DISSCHARGE
AND NOT   M00592	// HOLD DISSCHARGE
MPUSH
AND NOT   M0001F	// M_HIGH UNDERHOPER PACKER
AND NOT   M00023	// KUNCI MIXER OPEN
AND NOT   M0080D	// START CLOSE DOOR 
AND NOT   T0025	// TIMER KUNCI OPEN DOOR
OUT       M0080C	// START OPEN DOOR 
MLOAD
LOAD      M0001D	// M_SENSOR OPEN DOOR MIXER 
OR        M00023	// KUNCI MIXER OPEN
AND LOAD
OUT       M0070C	// DISSCHARGE MIXER 
TON       T0025 25	// TIMER KUNCI OPEN DOOR
MPUSH
AND       M0070C	// DISSCHARGE MIXER 
ANDP      F00093
AND NOT   M0080E	// STOP UNDERHOPPER PROSES
ADD       D00153 1 D00153	// COUNTING DISSCHARGE / COUNTING DISSCHARGE
MPOP
AND>=     D00153 30	// COUNTING DISSCHARGE
OUT       M0080E	// STOP UNDERHOPPER PROSES
MLOAD
AND       M0080E	// STOP UNDERHOPPER PROSES
OUT       M00415	// AUTO_SCADA21 AUTO CLOSE DOOR MIXER 
MPOP
AND       M00415	// AUTO_SCADA21 AUTO CLOSE DOOR MIXER 
AND       M0001E	// M_SENSOR CLOSE DOOR MIXER
TON       T0021 150	// TIMER OFF DISSCHARGE MIXER
; L24
LOADP     T0021	// TIMER OFF DISSCHARGE MIXER
MOV       0 D00153	// COUNTING DISSCHARGE
; L25
LOADP     M0001D	// M_SENSOR OPEN DOOR MIXER 
OR        M00023	// KUNCI MIXER OPEN
AND NOT   T0021	// TIMER OFF DISSCHARGE MIXER
AND NOT   M00450	// RESET BATCH
OUT       M00023	// KUNCI MIXER OPEN
; L27
LOAD      F00099
MPUSH
AND       M00830	// START MIXING 
MOV       D00151 D01239	// COUNTING MIXER
MPOP
AND       M0080B	// PROSES UNDERHOPPER DISSCHARGE
MOV       D00153 D01239	// COUNTING DISSCHARGE
; L29
LOAD      F00099
AND NOT   M00830	// START MIXING 
AND NOT   M0080B	// PROSES UNDERHOPPER DISSCHARGE
MOV       0 D01239

PROGRAM ProsesRecord (task: Scan Program)

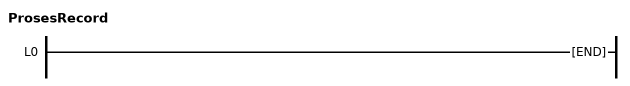
; L0
END

PROGRAM End (task: Scan Program)

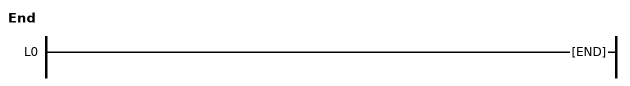
; L0
END

VARIABLES AND COMMENTS (devices not used above)
M00400	BIT	AUTO_SCADA // START AUTO PROSES 
M0040A	BIT	AUTO_SCADA10 // AUTO SCREW HOPPER JETFLO PASIR HALUS 
M0040C	BIT	AUTO_SCADA12 // AUTO SCREW HOPPER PASIR KASAR 
M00412	BIT	AUTO_SCADA18 // READY ADDITIF MIXER 
M00413	BIT	AUTO_SCADA19 // AUTO SAMPLE MIXER 
M00416	BIT	AUTO_SCADA22 // AUTO RUN MOTOR HIDROLIK MIXER 
M00417	BIT	AUTO_SCADA23 // HOLD TRANSFER
M00418	BIT	AUTO_SCADA24 // HOLD WEIGHING
M00419	BIT	AUTO_SCADA25 // HOLD DISSCHARGE MIXER 
M00407	BIT	AUTO_SCADA7 // AUTO SCREW HOPPER JETFLO POWDER
M00300	BIT	MEMORY_MANUAL // AUTO/MANUAL SCADA
M0030F	BIT	MEMORY_MANUAL15 // MANUAL JETFLO PASIR KASAR 02
M00316	BIT	MEMORY_MANUAL22 // MANUAL SAMPLE MIXER 
M00317	BIT	MEMORY_MANUAL23 // MANUAL START MIXER 
M00305	BIT	MEMORY_MANUAL5 // MANUAL SCREW EX GROUT SEMEN GREY 
M00306	BIT	MEMORY_MANUAL6 // MANUAL SCREW EX GROUT CALCITE
M00307	BIT	MEMORY_MANUAL7 // MANUAL SCREW HOPPER JETFLO POWDER 
M00308	BIT	MEMORY_MANUAL8 // MANUAL SCREW HOPPER JETFLO PASIR HALUS 
M00309	BIT	MEMORY_MANUAL9 // MANUAL SCREW HOPPER JETFLO PASIR KASAR 
P0002A	BIT	OUPTUT_10 // KONTAKTOR SCREW HOPPER PASIR
P00033	BIT	OUPTUT_19 // CHOPPER 01,02,03
P00038	BIT	OUPTUT_24 // SIRINE AUTO CYCLE TIME FEEDING POWDER
P00039	BIT	OUPTUT_25 // SIRINE AUTO CYCLE TIME FEEDING PASIR 
P0003A	BIT	OUPTUT_26 // LAMPU ADDITIF READY MIXER
P0003C	BIT	OUPTUT_28 // ZERO INDIKATOR POWDER
P0003D	BIT	OUPTUT_29 // TARE INDIKATOR POWDER
P0003E	BIT	OUPTUT_30 // SPARE
P0003F	BIT	OUPTUT_31 // SPARE
R00000	WORD	tmr10
D00010	WORD	DATA SEMEN
D00018	WORD	OFF VALVE SEMEN
D00020	WORD	DATA OFFSET SEMEN
D00022	WORD	TARGET SEMEN
D00024	WORD	OFF VALVE SEMEN
D00030	WORD	DATA KAPUR
D00038	WORD	OFFSET VALVE KAPUR
D00040	WORD	DATA OFFSET KAPUR
D00042	WORD	OFF VALVE KAPUR
D00044	WORD	TARGET KAPUR
D01000	WORD	DATA INDIKATOR 1
D01500	WORD	TARGET SEMEN + KAPUR
D01502	WORD	OFF VALVE SEMEN + KAPUR
D02000	WORD	Serial PC
D02021	WORD	Serial PC Save02
P00100	BIT	SELECTAUTO
P00101	BIT	SELECTMANUAL
D00100	WORD	TARGET SEMEN
D00101	WORD	TARGET KAPUR
D00102	WORD	TARGET SEMEN PUTIH
D00103	WORD	TARGET PASIR
M00032	BIT	M_RECORD HASIL SEMEN
D00104	WORD	TARGET SEMEN PUTIH
M00034	BIT	M_RECORD HASIL KAPUR
T0101	BIT/WORD	WaktuMixing
T0102	BIT/WORD	T_SelesaiMix
D00200	WORD	FINE SEMEN
D00201	WORD	FINE KAPUR
D00203	WORD	FINE SEMEN  PUTIH
D00202	WORD	FINE PASIR
D00304	WORD	HASIL FINE SEMEN PUTIH
T0080	BIT/WORD	T_OFF RECORD PASIR KASAR
M00059	BIT	M_RECORD HASIL PASIR KASAR
T0040	BIT/WORD	T_START FILLING SEMEN PUTIH
M00900	BIT	BatchPindah
D01100	WORD	DATA INDIKATOR 2
K0100	WORD	SET FRQ
D02600	WORD	OUTPUT INV
D02601	WORD	CMD01
M00117	BIT	START HIGH INV SC ABU
M00118	BIT	START LOW INV SC ABU
M00119	BIT	STOP RUN INV SCREW
M0011A	BIT	MEMORI FOR RUN INV SC01
M0011B	BIT	MEMORI REV RUN INV SC01
M00127	BIT	START HIGH INV SC KAPUR
M00128	BIT	START LOW INV SC KAPUR
M00137	BIT	START HIGH INV SC KASAR
M00138	BIT	START LOW INV SC KASAR
M00147	BIT	START HIGH INV SC HALUS
M00148	BIT	START LOW INV SC HALUS
D01050	WORD	DATA TIMBANGAN HOPPER
D01150	WORD	DATA TIMBANGAN PACKER
D03010	WORD	HASIL SEMEN PUTIH
D03040	WORD	HASIL PASIR HALUS
D03000	WORD	HASIL SEMEN ABU2
D03004	WORD	TARGET ABU+KAPUR
D03022	WORD	HASIL KAPUR-ABU
D03024	WORD	HASIL KAPUR-PUTIH
D03026	WORD	TARGET ABU+KAPUR+KASAR
D03028	WORD	TARGET PUTIH+KAPUR+KASAR
D03032	WORD	HASIL KASAR-KAPUR-ABU
D03034	WORD	HASIL KASAR-KAPUR-PUTIH
D03036	WORD	TARGET HALUS+KAPUR+ABU
D03038	WORD	TARGET HALUS+KAPUR+PUTIH
D03050	WORD	HASIL KAPUR
D03020	WORD	SWEP HASIL KAPUR
D03030	WORD	SWEP HASIL PASIR KASAR
D03060	WORD	HASIL PASIR KASAR
D03070	WORD	HASIL PASIR HALUS
M02110	BIT	START JETFLO
M02124	BIT	START KAPUR
M02126	BIT	START KASAR
M02128	BIT	START HALUS
M00122	BIT	SELASAI MIXING
D00318	WORD	HASIL TOTAL FORMULA
D00305	WORD	HASIL FINE ADITIF
D03084	WORD	TARGET HASIL ADITIF+PUTIH+KAPUR+PASIR
D03082	WORD	TARGET HASIL ADITIF+ABU+KAPUR+PASIR
D03090	WORD	HASIL ADITIF 
M0212A	BIT	START ADITIF
K3400	WORD	TARGET SEMEN ABU
D00110	WORD	TARGET KURANG SEMEN PUTIH
K3402	WORD	OFFSET SEMEN ABU
D00120	WORD	OFFSET SEMEN ABU
K3404	WORD	FINE SEMEN ABU
D00130	WORD	FINE SEMEN ABU
K3406	WORD	TARGET VIBRO 
D00140	WORD	TARGET VIBRO
M02120	BIT	START HIGH ABU
M00150	BIT	START LOW ABU
D00310	WORD	FINE KAPUR
D00320	WORD	FINE KASAR
D00322	WORD	CORSE KASAR
D00330	WORD	FINE HALUS
D00332	WORD	CORSE HALUS
D00340	WORD	FINE ADITIF
D00350	WORD	FINE PUTIH
D00352	WORD	CORSE PUTIH
D00342	WORD	CORSE ADITIF
M00152	BIT	FINISH ABU
M02130	BIT	START HIGH KAPUR
M00160	BIT	START LOW KAPUR
T0071	BIT/WORD	TON KAPUR
T0072	BIT/WORD	TON KASAR
T0070	BIT/WORD	TON ABU
M02140	BIT	START HIGH KASAR
M00172	BIT	FINISH KASAR
M00170	BIT	START LOW KASAR
T0073	BIT/WORD	TON HALUS
M00182	BIT	FINISH HALUS
M00180	BIT	START LOW HALUS
M02150	BIT	START HIGH HALUS
T0074	BIT/WORD	TON PUTIH
M02160	BIT	START HIGH PUTIH
M00190	BIT	START LOW PUTIH
M00192	BIT	FINISH PUTIH
T0075	BIT/WORD	TON ADITIF
M02200	BIT	START HIGH ADITIF
M02004	BIT	ISI ADITIF
M00080	BIT	M START AUTO
T0050	BIT/WORD	T SIMPAN ABU
T0060	BIT/WORD	T RESET ABU
M00020	BIT	ABU
M00022	BIT	KAPUR
M00024	BIT	KASAR
M00026	BIT	HALUS
M00028	BIT	PUTIH
M0002A	BIT	ADITIF
M00200	BIT	START LOW ADITIF
M00202	BIT	FINISH ADITIF
M00162	BIT	FINISH KAPUR
D00314	WORD	FINE KAPUR
D00316	WORD	CORSE KAPUR
D03210	WORD	SWEP KAPUR
D00324	WORD	FINE KASAR
D00326	WORD	CORSE KASAR
D00334	WORD	FINE HALUS
D00336	WORD	CORSE HALUS
D03230	WORD	SWEP HALUS
D03220	WORD	SWEP KASAR
D03080	WORD	HASIL SEMEN PUITH
D03240	WORD	SWEP PUTIH
D03100	WORD	HASIL ADITIF
T0062	BIT/WORD	SIMPAN KAPUR
T0052	BIT/WORD	SIMPAN SWEP KAPUR
T0053	BIT/WORD	SIMPAN SWEP KASAR
T0063	BIT/WORD	SIMPAN KASAR
T0054	BIT/WORD	SIMPAN SWEP HALUS
T0064	BIT/WORD	SIMPAN HALUS
T0051	BIT/WORD	SIMPAN SWEP PUTIH
T0061	BIT/WORD	SIMPAN PUTIH
T0065	BIT/WORD	SIMPAN ADITIF
T0076	BIT/WORD	START MIXER
D00354	WORD	FINE PUTIH
D00356	WORD	CORSE PUTIH
T0092	BIT/WORD	T FINISH KASAR
T0093	BIT/WORD	T FINISH HALUS
T0091	BIT/WORD	T FINISH KAPUR
T0094	BIT/WORD	T FINISH PUTIH
T0095	BIT/WORD	T FINISH ADITIF
T0077	BIT/WORD	FINISH PENIMBANGAN
D03200	WORD	SWEP ABU
T0082	BIT/WORD	T KAPUR
T0083	BIT/WORD	T KASAR
T0084	BIT/WORD	T HALUS
T0081	BIT/WORD	T PUTIH
T0085	BIT/WORD	T ADITIF
T0090	BIT/WORD	FINISH ABU
M00092	BIT	ZERO
M00090	BIT	PENIMBANGAN FINISH
M00130	BIT	FINISH BATCH
K0030	WORD	COUNTER TIMBANG
K0040	WORD	COUNTER BATCH
M00100	BIT	MIX TIME
T0106	BIT/WORD	T OFF MIXER
T0105	BIT/WORD	T DOOR CLOSE
M00110	BIT	OPEN TIMBANGAN
T0089	BIT/WORD	T CLOSE TIMBANGAN
M02010	BIT	SIM ABU
M02011	BIT	SIM KAPUR
M02012	BIT	SIM KASAR
M02013	BIT	SIM HALUS
M02014	BIT	SIM PUTIH
M02015	BIT	SIM ADITIF
M02020	BIT	TIME SQUEN
M02022	BIT	TIME RECORD
T0100	BIT/WORD	T OPEN TIMBANGAN
T0097	BIT/WORD	START SQUEN TIMBANG
T0088	BIT/WORD	AUTO ZERO
M00095	BIT	M ADITIF ISI
D00080	WORD	HOPPER FULL
M00132	BIT	FINISH TIMBANG
K0035	WORD	COUNTER MIXING
M00107	BIT	COUNTER MIXING
M00133	BIT	FINISH MIXER
M00210	BIT	M FINISH TIMBANG
T0098	BIT/WORD	START SQUEN MIXER
T0110	BIT/WORD	START SQUEN FULL
D00410	WORD	Hasil2
D00420	WORD	Hasil3
D00430	WORD	Hasil4
D00440	WORD	Total
M00157	BIT	START HIGH INV SC PUTIH
M00158	BIT	START LOW INV SC PUTIH
M00049	BIT	ANGKA TIMBANGAN
M00125	BIT	M CLOSE TIMBANGAN
M00490	BIT	SQUEN FINISH PENIMBANGAN
M00094	BIT	HOLD TIMBANG
M00123	BIT	OPEN MIXER
K0045	WORD	LOCK FINISH TIMBANG
M02006	BIT	PB FULL HOPPER
K0050	WORD	LOCK FINISH MIXING
M02001	BIT	PB HMI STOP AUTO 
M02000	BIT	PB HMI START AUTO
M02003	BIT	PB HMI HOLD TIMBANG
M02005	BIT	PB HMI HOLD MIXER
M00135	BIT	PB HMI HOPPER FULL
M00070	BIT	M_RECORD HASIL SEMEN PUTIH
M00035	BIT	M_START MIXER
M00060	BIT	M_RECORD HASIL PASIR HALUS
M00075	BIT	M_RECORD HASIL ADITIF
M00105	BIT	COUNTER TIMBANG
M00102	BIT	COUNTER BATCH
M02008	BIT	PB HMI START MIXER
K0110	WORD	TON ABU
K0112	WORD	FINISH ABU
K0114	WORD	TON KAPUR
K0116	WORD	FINISH KAPUR
K0118	WORD	TON KASAR
K0120	WORD	FINISH KASAR
K0122	WORD	TON HALUS
K0124	WORD	FINISH HALUS
K0126	WORD	TON PUTIH
K0128	WORD	FINISH PUTIH
K0130	WORD	TON ADITIF
K0132	WORD	FINISH ADITIF
K0134	WORD	TON MIXER
K0136	WORD	FINISH TIMBANG
K0200	WORD	T RECORD ABU
K0202	WORD	T RECORD KAPUR
K0204	WORD	T RECORD KASAR
K0206	WORD	T RECORD HALUS
K0208	WORD	T RECORD PUTIH
K0210	WORD	T RECORD ADITIF
K0220	WORD	T OPEN TIMBANG
K0222	WORD	T CLOSE TIMBANG
K0224	WORD	T AUTO ZERO
K0226	WORD	T CLOSE DOOR
K0230	WORD	T START SQUEN
K0240	WORD	MIXING TIME
K1160	WORD	H FRQ KAPUR
K1170	WORD	H FRQ KASAR
K1180	WORD	H FRQ HALUS
K1190	WORD	H FRQ PUTIH
K1152	WORD	L FRQ ABU
K1162	WORD	L FRQ KAPUR
K1172	WORD	L FRQ KASAR
K1182	WORD	L FRQ HALUS
K1192	WORD	L FRQ PUTIH
D03250	WORD	SWEP ADTIF
K0150	WORD	LOCK RECORD ABU
K0152	WORD	LOCK  RECORD KAPUR
K0154	WORD	LOCK RECORD KASAR
K0156	WORD	LOCK RECORD HALUS
K0158	WORD	LOCK RECORD PUTIH
K0160	WORD	LOCK RECORD ADITIF
M0002F	BIT	LAMPU MIXING
K3350	WORD	SIMULATOR TIMBANGAN
K3355	WORD	TARGET PACKER
K0025	WORD	TARGET PRODUKSI
K3360	WORD	DISPLAY MIXING
M00082	BIT	M START MANUAL
D00344	WORD	FINE ADITIF
D00346	WORD	CORSE ADITIF
M0007A	BIT	M_RECORD ALL PENIMBANGAN
M00085	BIT	M START AUTO SQUEN
T0112	BIT/WORD	T OFF SQUEN TIMBANG
T0131	BIT/WORD	T RESET PUTIH
T0132	BIT/WORD	T RESET KAPUR
T0133	BIT/WORD	T RESET KASAR
T0134	BIT/WORD	T RESET HALUS
T0135	BIT/WORD	T RESET ADITIF
M00136	BIT	M FULL HOPPER
D00714	WORD	TARGET OFF PACKER
D00712	WORD	TARGET FINE
D00710	WORD	FINE AUTO
T0150	BIT/WORD	T SIMPAN PACKER
T0151	BIT/WORD	T START CORRECTION
T0152	BIT/WORD	T LOCK CORRECTION
K0250	WORD	SET CORRECTION PACKER
K0248	WORD	SET FINE PACKER
M00270	BIT	TEST OL INVERTER
D00406	WORD	HSP1
D00416	WORD	HSP2
D00426	WORD	HSP3
D00436	WORD	HSP4
D00446	WORD	TOTAL HASIL PENIMBANGAN
D00412	WORD	HST2
D00422	WORD	HST3
D00432	WORD	HST4
D00444	WORD	TOTAL HASIL TARGET
M01250	BIT	M RECORD HMI
M0011D	BIT	MEMORI OL INVERTER SC
M0010C	BIT	start mixing time
M00120	BIT	COUNTING MIXING
K0060	WORD	LOCK CORRECTION
M00250	BIT	M START SIMPAN PACKER
M00252	BIT	M SIMPAN +
M00254	BIT	M SIMPAN -
M00256	BIT	M BATAS ZERO
M0010A	BIT	M COUTING TOMBOL MIXER
K0070	WORD	on vibro
K0072	WORD	off vibro
K0074	WORD	on vibro kapur
K0076	WORD	off vibro kapur
D00800	WORD	data scanner
K3365	WORD	counting pb manual
K0170	WORD	LOCK COUNTING TIMBANG
T0170	BIT/WORD	T LOCK COUNTING TIMBANG
K0047	WORD	LOCK COUNTING MIXING
K0182	WORD	LOCK TARGET KAPUR
K0184	WORD	LOCK TARGET KASAR
K0186	WORD	LOCK TARGET HALUS
K0188	WORD	LOCK TARGET PUTIH
K0190	WORD	LOCK TARGET ADITIF
K0180	WORD	LOCK TARGET ABU
T0160	BIT/WORD	TON VIBRO WH
T0162	BIT/WORD	TOFF VIBRO WH
T0164	BIT/WORD	TON VIBRO KAPUR
T0166	BIT/WORD	TOFF VIBRO KAPUR
K0003	WORD	MAXIMAL SEMEN ABU SCADA
K0004	WORD	MINIMAL SEMEN ABU SCADA
D00312	WORD	HASIL MINIMAL SEMEN ABU PLC
K0008	WORD	MAXIMAL SEMEN PUTIH SCADA
K0009	WORD	MINIMAL SEMEN PUTIH SCADA
K0013	WORD	MAXIMAL KAPUR SCADA
K0014	WORD	MINIMAL KAPUR SCADA
K0018	WORD	MAXIMAL PASIR KASAR SCADA
K0019	WORD	MINIMAL PASIR KASAR SCADA
K0023	WORD	MAXIMAL PASIR HALUS SCADA
K0024	WORD	MINIMAL PASIR HALUS SCADA
M0001C	BIT	M_OL CHOPPER 03
M0031A	BIT	MANUAL VIBRO MOTOR SEMEN GREY 
M0031B	BIT	MANUAL VIBRO MOTOR CALCITE
M00500	BIT	START ADDITIF
M00501	BIT	FINISH ADDITIF 
M00502	BIT	STOP ADDITIF 
M00503	BIT	RESET ADDITIF 
M00505	BIT	PROSES TIMBANG ADDITIF 
D00263	WORD	HASIL A DAN B ADDITIF
D00264	WORD	HASIL C DAN D ADDITIF
D00265	WORD	HASIL E DAN F ADDITIF
D00266	WORD	HASIL G DAN H ADDITIF
D00268	WORD	HASIL ABCD
D00269	WORD	HASIL EFGH
D00271	WORD	FINISH HASIL ADDITIF
M00605	BIT	STOP TIMER SEMEN GREY 
M00607	BIT	STOP SEMI MANUAL SEMEN GREY
M00611	BIT	STOP TIMER KAPUR
M00613	BIT	STOP SEMI MANUAL KAPUR
M0061D	BIT	STOP TIMER SEMEN PUTIH
M0061F	BIT	STOP SEMI MANUAL SEMEN PUTIH
M00620	BIT	START BV SCREW SEMEN PUTIH
D00006	WORD	SIMPAN INDIKATOR PASIR KASAR
D00007	WORD	SIMPAN INDIKATOR PASIR HALUS
D00111	WORD	TARGET KURANG PASIR KASAR
D00112	WORD	TARGET KURANG PASIR HALUS
M00629	BIT	STOP TIMER PASIR  KASAR
M0062B	BIT	STOP SEMI MANUAL PASIR KASAR
M0062C	BIT	START BV SCREW PASIR KASAR
M00635	BIT	STOP TIMER PASIR   HALUS
M00637	BIT	STOP SEMI MANUAL PASIR  HALUS
M00638	BIT	START BV SCREW PASIR  HALUS
M00801	BIT	STOP PROSES MATERIAL 
T0019	BIT/WORD	TIMER OFF HOPPER PASIR 
M0080A	BIT	STOP UNDERHOPPER PROSES
D00152	WORD	TIMER DISCCHARGE
K1140	WORD	HIGH SEMEN PUTIH 
K1141	WORD	LOW SEMEN PUTIH 
M00710	BIT	RVS POWDER
M00596	BIT	BYPAS ADD
D00275	WORD	ACTUAL ADDITIF A
D00276	WORD	ACTUAL ADDITIF B
D00277	WORD	ACTUAL ADDITIF C
D00278	WORD	ACTUAL ADDITIF D
D00279	WORD	ACTUAL ADDITIF E
D00280	WORD	ACTUAL ADDITIF F
D00281	WORD	ACTUAL ADDITIF G
D00282	WORD	ACTUAL ADDITIF H
M00640	BIT	READY PRINT ADDA
M00641	BIT	READY PRINT ADD B
M00643	BIT	READY PRINT ADD D
M00642	BIT	READY PRINT ADDITIF C
D00175	WORD	ACTUAL SEMEN PUTIH
M00354	BIT	PERBARUI INDIKATOR
M00680	BIT	DOSS ERROR
K0261	WORD	DRIBBLE KAPUR SCADA
K0532	WORD	DRIBBLE PASIR KASAR SCADA